(****************************************************************************************************<br>
© Syntegon Group.<br>
All rights reserved, also regarding any disposal, exploitation, reproduction, editing, distribution,<br>
as well as in the event of applications for industrial property rights.<br>
*****************************************************************************************************<br>
DESCRIPTION:<br>
Answers the waiting machine command: accepted, or rejected with the reason the Simulator shows. The command no<br>
longer waits afterwards.<br>
*****************************************************************************************************<br>
OUTPUT VALUES:<br>
FALSE while no command waits.<br>
****************************************************************************************************)
METHOD m_AnswerCommand : BOOL
VAR_INPUT
	vi_b_Accepted						: BOOL;	// TRUE: the application carries the command out
	vi_str_Reason						: STRING(80);	// why it is rejected, '' when accepted
END_VAR
m_AnswerCommand := vo_Config.stCommand.bRequested;
IF NOT m_AnswerCommand THEN
	RETURN;
END_IF
vo_Config.stCommandStatus.nHandledCommandId := vo_Config.stCommand.nCommandId;
vo_Config.stCommandStatus.eResult := SEL(vi_b_Accepted, E_ConfigCommandResult.REJECTED, E_ConfigCommandResult.ACCEPTED);
vo_Config.stCommandStatus.sMessage := SEL(vi_b_Accepted, vi_str_Reason, '');
vo_Config.stCommand.bRequested := FALSE;
END_METHOD

(****************************************************************************************************<br>
© Syntegon Group.<br>
All rights reserved, also regarding any disposal, exploitation, reproduction, editing, distribution,<br>
as well as in the event of applications for industrial property rights.<br>
*****************************************************************************************************<br>
DESCRIPTION:<br>
The machine command waiting for the application's answer (START, STOP, RESET); NONE while none waits. Answer it<br>
with m_AnswerCommand: the application alone decides whether it is carried out.<br>
****************************************************************************************************)
METHOD m_Command : E_ConfigCommand
IF vo_Config.stCommand.bRequested THEN
	m_Command := vo_Config.stCommand.eCommand;
ELSE
	m_Command := E_ConfigCommand.NONE;
END_IF
END_METHOD

(****************************************************************************************************<br>
© Syntegon Group.<br>
All rights reserved, also regarding any disposal, exploitation, reproduction, editing, distribution,<br>
as well as in the event of applications for industrial property rights.<br>
*****************************************************************************************************<br>
DESCRIPTION:<br>
Every cycle, after the fields are declared: handles a staged recipe or a reset (a recipe only while<br>
vi_b_ApplyAllowed), keeps the active recipe in vio_Set and gives the effective values in vo_Config.aActive: the<br>
active recipe while one is valid, else the fields' program values.<br>
*****************************************************************************************************<br>
OUTPUT VALUES:<br>
TRUE in the cycle a recipe was taken over or reset.<br>
****************************************************************************************************)
METHOD m_Cycle : BOOL
VAR_IN_OUT
	vio_Set								: ST_ConfigRecipeSet;	// the application's VAR PERSISTENT active recipe
END_VAR
VAR_INPUT
	vi_b_ApplyAllowed					: BOOL;	// [-] a staged recipe may be taken over now, e.g. while the machine stands
END_VAR
VAR
	str_TempRejection					: STRING(80);
	un_TempIndex						: UINT;
END_VAR
m_Cycle := FALSE;
CASE m_Staging(vio_Staging := vo_Config.stStaging, vio_Status := vo_Config.stStatus, vi_b_ApplyAllowed := vi_b_ApplyAllowed,
	vi_udn_ActiveVersion := SEL(vio_Set.bValid, 0, vio_Set.nVersion)) OF
	E_ConfigAction.RESET:
		vio_Set.bValid := FALSE;
		m_Handled(vio_Staging := vo_Config.stStaging, vio_Status := vo_Config.stStatus, vi_str_Rejection := '');
		m_Cycle := TRUE;
	E_ConfigAction.TAKE_OVER:
		str_TempRejection := m_Invalid();
		IF str_TempRejection = '' THEN
			vio_Set.nLastVersion := vio_Set.nLastVersion + 1;
			vio_Set.nVersion := vio_Set.nLastVersion;
			vio_Set.aValues := vo_Config.aStaged;
			vio_Set.bValid := TRUE;
			m_Cycle := TRUE;
		END_IF
		m_Handled(vio_Staging := vo_Config.stStaging, vio_Status := vo_Config.stStatus, vi_str_Rejection := str_TempRejection);
END_CASE


(****************************************************************************************************
EFFECTIVE VALUES
****************************************************************************************************)
un_TempIndex := 0;
WHILE un_TempIndex < vo_Config.nFieldCount AND un_TempIndex < CONFIG_GlobalConst_Param.CONFIG_un_MAX_RECIPE_FIELDS DO
	vo_Config.aActive[un_TempIndex] := SEL(vio_Set.bValid, vo_Config.aFields[un_TempIndex].fProgramValue,
		vio_Set.aValues[un_TempIndex]);
	un_TempIndex := un_TempIndex + 1;
END_WHILE
vo_Config.stStatus.nActiveVersion := SEL(vio_Set.bValid, 0, vio_Set.nVersion);
END_METHOD

(****************************************************************************************************<br>
© Syntegon Group.<br>
All rights reserved, also regarding any disposal, exploitation, reproduction, editing, distribution,<br>
as well as in the event of applications for industrial property rights.<br>
*****************************************************************************************************<br>
DESCRIPTION:<br>
Declares recipe field vi_un_Field (1..CONFIG_un_MAX_RECIPE_FIELDS): its name, the component it belongs to, how its<br>
value is kept, its unit, range and the program value that applies while no recipe is active. Fields are listed up<br>
to the highest one declared. Idempotent: call it every cycle, before m_Cycle. A CHOICE field's values are named with<br>
m_SetChoice and range from 0; its vi_lr_Min and vi_lr_Max are not used, nor a SWITCH's.<br>
*****************************************************************************************************<br>
OUTPUT VALUES:<br>
FALSE for vi_un_Field = 0 or above CONFIG_un_MAX_RECIPE_FIELDS.<br>
****************************************************************************************************)
METHOD m_DeclareField : BOOL
VAR_INPUT
	vi_un_Field							: UINT;	// [-] 1..CONFIG_un_MAX_RECIPE_FIELDS
	vi_str_Name							: STRING(31);	// unique in the recipe, e.g. 'BeltSpeed'
	vi_udn_Group						: UDINT;	// [-] manifest id of the Syn_Visu component, 0 = the whole machine
	vi_e_Type							: E_ConfigFieldType;
	vi_str_Unit							: STRING(15);	// e.g. 'mm/s', '' = none
	vi_lr_Min							: LREAL;	// smallest value of a NUMBER or INTEGER field
	vi_lr_Max							: LREAL;	// largest value of a NUMBER or INTEGER field
	vi_lr_ProgramValue					: LREAL;	// the application's own value; a SWITCH: 1 = on
END_VAR
m_DeclareField := vi_un_Field > 0 AND vi_un_Field <= CONFIG_GlobalConst_Param.CONFIG_un_MAX_RECIPE_FIELDS;
IF NOT m_DeclareField THEN
	RETURN;
END_IF
vo_Config.aFields[vi_un_Field - 1].sName := vi_str_Name;
vo_Config.aFields[vi_un_Field - 1].nGroup := vi_udn_Group;
vo_Config.aFields[vi_un_Field - 1].eType := vi_e_Type;
vo_Config.aFields[vi_un_Field - 1].sUnit := vi_str_Unit;
vo_Config.aFields[vi_un_Field - 1].fMin := vi_lr_Min;
vo_Config.aFields[vi_un_Field - 1].fMax := vi_lr_Max;
vo_Config.aFields[vi_un_Field - 1].fProgramValue := vi_lr_ProgramValue;
IF vi_un_Field > vo_Config.nFieldCount THEN
	vo_Config.nFieldCount := vi_un_Field;
END_IF
END_METHOD

(****************************************************************************************************<br>
© Syntegon Group.<br>
All rights reserved, also regarding any disposal, exploitation, reproduction, editing, distribution,<br>
as well as in the event of applications for industrial property rights.<br>
*****************************************************************************************************<br>
DESCRIPTION:<br>
Effective value of an INTEGER or CHOICE recipe field as a whole number (see m_Value).<br>
****************************************************************************************************)
METHOD m_Integer : DINT
VAR_INPUT
	vi_un_Field							: UINT;	// [-] 1..the field count
END_VAR
m_Integer := LREAL_TO_DINT(m_Value(vi_un_Field := vi_un_Field));
END_METHOD

(****************************************************************************************************<br>
© Syntegon Group.<br>
All rights reserved, also regarding any disposal, exploitation, reproduction, editing, distribution,<br>
as well as in the event of applications for industrial property rights.<br>
*****************************************************************************************************<br>
DESCRIPTION:<br>
Why the staged recipe cannot be taken over; '' when it can: a value outside its field's range (NUMBER, INTEGER),<br>
not one of its choices (CHOICE), not a whole number (INTEGER, CHOICE) or not 0 or 1 (SWITCH).<br>
****************************************************************************************************)
METHOD PRIVATE m_Invalid : STRING(80)
VAR
	un_TempIndex						: UINT;
	lr_TempValue						: LREAL;
	lr_TempMin							: LREAL;
	lr_TempMax							: LREAL;
END_VAR
m_Invalid := '';
un_TempIndex := 0;
WHILE un_TempIndex < vo_Config.nFieldCount AND un_TempIndex < CONFIG_GlobalConst_Param.CONFIG_un_MAX_RECIPE_FIELDS DO
	lr_TempValue := vo_Config.aStaged[un_TempIndex];
	CASE vo_Config.aFields[un_TempIndex].eType OF
		E_ConfigFieldType.SWITCH:
			lr_TempMin := 0;
			lr_TempMax := 1;
		E_ConfigFieldType.CHOICE:
			lr_TempMin := 0;
			lr_TempMax := UINT_TO_LREAL(vo_Config.aFields[un_TempIndex].nChoiceCount) - 1;
	ELSE
		lr_TempMin := vo_Config.aFields[un_TempIndex].fMin;
		lr_TempMax := vo_Config.aFields[un_TempIndex].fMax;
	END_CASE
	(* The range first: only a value in range is turned into a whole number. NaN equals nothing, not even itself. *)
	IF lr_TempValue <> lr_TempValue OR lr_TempValue < lr_TempMin OR lr_TempValue > lr_TempMax THEN
		m_Invalid := CONCAT(CONCAT('Field ', vo_Config.aFields[un_TempIndex].sName), CONCAT(': ', CONCAT(LREAL_TO_STRING(lr_TempValue),
			CONCAT(' is outside ', CONCAT(LREAL_TO_STRING(lr_TempMin), CONCAT(' to ', LREAL_TO_STRING(lr_TempMax)))))));
		RETURN;
	END_IF
	IF vo_Config.aFields[un_TempIndex].eType <> E_ConfigFieldType.NUMBER
		AND LINT_TO_LREAL(LREAL_TO_LINT(lr_TempValue)) <> lr_TempValue
	THEN
		m_Invalid := CONCAT(CONCAT('Field ', vo_Config.aFields[un_TempIndex].sName), CONCAT(': ',
			CONCAT(LREAL_TO_STRING(lr_TempValue), ' is not a value of its type')));
		RETURN;
	END_IF
	un_TempIndex := un_TempIndex + 1;
END_WHILE
END_METHOD

(****************************************************************************************************<br>
© Syntegon Group.<br>
All rights reserved, also regarding any disposal, exploitation, reproduction, editing, distribution,<br>
as well as in the event of applications for industrial property rights.<br>
*****************************************************************************************************<br>
DESCRIPTION:<br>
Names value vi_un_Value (0..CONFIG_un_MAX_CHOICES-1) of the CHOICE field vi_un_Field, e.g. 0 = 'Lanes'. The field<br>
has as many choices as the highest value named plus one. Idempotent: call it every cycle with m_DeclareField.<br>
*****************************************************************************************************<br>
OUTPUT VALUES:<br>
FALSE for a field not declared or a value above CONFIG_un_MAX_CHOICES - 1.<br>
****************************************************************************************************)
METHOD m_SetChoice : BOOL
VAR_INPUT
	vi_un_Field							: UINT;	// [-] the field, 1..its count
	vi_un_Value							: UINT;	// [-] the value it names, from 0
	vi_str_Text							: STRING(31);	// e.g. 'Lanes'
END_VAR
m_SetChoice := vi_un_Field > 0 AND vi_un_Field <= vo_Config.nFieldCount
	AND vi_un_Value < CONFIG_GlobalConst_Param.CONFIG_un_MAX_CHOICES;
IF NOT m_SetChoice THEN
	RETURN;
END_IF
vo_Config.aFields[vi_un_Field - 1].aChoices[vi_un_Value] := vi_str_Text;
IF vi_un_Value >= vo_Config.aFields[vi_un_Field - 1].nChoiceCount THEN
	vo_Config.aFields[vi_un_Field - 1].nChoiceCount := vi_un_Value + 1;
END_IF
END_METHOD

(****************************************************************************************************<br>
© Syntegon Group.<br>
All rights reserved, also regarding any disposal, exploitation, reproduction, editing, distribution,<br>
as well as in the event of applications for industrial property rights.<br>
*****************************************************************************************************<br>
DESCRIPTION:<br>
Gives the declared field vi_un_Field the label the Simulator shows instead of its name put into words, and a<br>
description of what it is for, shown in the field's tooltip (config protocol 4, #49). Free text in the operators'<br>
language; the name stays the field's key. Idempotent: call it every cycle with m_DeclareField.<br>
*****************************************************************************************************<br>
OUTPUT VALUES:<br>
FALSE for a field not declared.<br>
****************************************************************************************************)
METHOD m_SetText : BOOL
VAR_INPUT
	vi_un_Field							: UINT;	// [-] the field, 1..its count
	vi_str_Label						: STRING(40);	// e.g. 'Belt speed', '' = the name put into words
	vi_str_Description					: STRING(160);	// what the field is for, '' = none
END_VAR
m_SetText := vi_un_Field > 0 AND vi_un_Field <= vo_Config.nFieldCount;
IF NOT m_SetText THEN
	RETURN;
END_IF
vo_Config.aFields[vi_un_Field - 1].sLabel := vi_str_Label;
vo_Config.aFields[vi_un_Field - 1].sDescription := vi_str_Description;
END_METHOD

(****************************************************************************************************<br>
© Syntegon Group.<br>
All rights reserved, also regarding any disposal, exploitation, reproduction, editing, distribution,<br>
as well as in the event of applications for industrial property rights.<br>
*****************************************************************************************************<br>
DESCRIPTION:<br>
Shows the declared field vi_un_Field in the Simulator only while field vi_un_OnField has the value vi_dn_Value<br>
(config protocol 4, #49), e.g. a lane count only while the pattern is Lanes. vi_un_OnField must be a SWITCH (0 / 1),<br>
CHOICE or INTEGER field and may belong to another group; a field depending on a hidden one is hidden too. A hidden<br>
field keeps its value and is written with the recipe. vi_un_OnField = 0 shows the field always. The gateway reports<br>
a condition on a NUMBER field, on the field itself, on a field not declared, on a value that field can never have<br>
or in a ring as a discovery error and shows that field always. Idempotent: call it every cycle with m_DeclareField.<br>
*****************************************************************************************************<br>
OUTPUT VALUES:<br>
FALSE for a field not declared.<br>
****************************************************************************************************)
METHOD m_SetVisibleWhen : BOOL
VAR_INPUT
	vi_un_Field							: UINT;	// [-] the field shown on condition, 1..its count
	vi_un_OnField						: UINT;	// [-] the field the condition reads, 0 = always shown
	vi_dn_Value							: DINT;	// [-] the value vi_un_OnField must have
END_VAR
m_SetVisibleWhen := vi_un_Field > 0 AND vi_un_Field <= vo_Config.nFieldCount;
IF NOT m_SetVisibleWhen THEN
	RETURN;
END_IF
vo_Config.aFields[vi_un_Field - 1].nVisibleField := vi_un_OnField;
vo_Config.aFields[vi_un_Field - 1].nVisibleValue := vi_dn_Value;
END_METHOD

(****************************************************************************************************<br>
© Syntegon Group.<br>
All rights reserved, also regarding any disposal, exploitation, reproduction, editing, distribution,<br>
as well as in the event of applications for industrial property rights.<br>
*****************************************************************************************************<br>
DESCRIPTION:<br>
Effective value of a SWITCH recipe field: TRUE for on (see m_Value).<br>
****************************************************************************************************)
METHOD m_Switch : BOOL
VAR_INPUT
	vi_un_Field							: UINT;	// [-] 1..the field count
END_VAR
m_Switch := m_Value(vi_un_Field := vi_un_Field) <> 0;
END_METHOD

(****************************************************************************************************<br>
© Syntegon Group.<br>
All rights reserved, also regarding any disposal, exploitation, reproduction, editing, distribution,<br>
as well as in the event of applications for industrial property rights.<br>
*****************************************************************************************************<br>
DESCRIPTION:<br>
Effective value of recipe field vi_un_Field, for the application's logic: the active recipe's, else the program<br>
value. 0 for a field not declared. A SWITCH gives 1 or 0, an INTEGER or CHOICE a whole number (m_Switch,<br>
m_Integer give them typed).<br>
****************************************************************************************************)
METHOD m_Value : LREAL
VAR_INPUT
	vi_un_Field							: UINT;	// [-] 1..the field count
END_VAR
IF vi_un_Field > 0 AND vi_un_Field <= vo_Config.nFieldCount THEN
	m_Value := vo_Config.aActive[vi_un_Field - 1];
ELSE
	m_Value := 0;
END_IF
END_METHOD

END_FUNCTION_BLOCK

// POUs/_FB_ConfigCartesian
(****************************************************************************************************<br>
© Syntegon Group.<br>
All rights reserved, also regarding any disposal, exploitation, reproduction, editing, distribution,<br>
as well as in the event of applications for industrial property rights.<br>
*****************************************************************************************************<br>
DESCRIPTION:<br>
Parameter set of one Cartesian robot (ADR 0017): its pose, origin shift, zones, gripper fingers, limit area and<br>
TCP limit area, written by the configurator, taken over when the application allows it.<br>
Typical cycle:<br>
  fb_CartParam.m_Register(vio_Manifest := GVL_Config.stManifest, vi_udn_Id := fb_Cart.m_Id());<br>
  fb_CartParam.m_Cycle(vio_Default := CartDefault, vio_Set := CartSet, vi_b_ApplyAllowed := b_Stopped);<br>
  fb_Cart.m_Configure(vi_Pose := fb_CartParam.m_Pose(), vi_lr_XMin := 0, ...);<br>
  fb_CartParam.m_PassOn(vio_Visu := fb_Cart);<br>
The application's logic takes its zones and limit areas from m_Active, not from its own constants.<br>
*****************************************************************************************************<br>
OUTPUT VALUES:<br>
vo_Config is the contract structure the gateway reads and writes at the path in the config manifest.<br>
*****************************************************************************************************<br>
VERSION         ¦ DATE       ¦ NAME      ¦ CHANGE<br>
Syn_Config 1.1.0 ¦ 2026-11-10 ¦ J.Willner ¦ New<br>
Syn_Config 2.0.0 ¦ 2026-11-11 ¦ J.Willner ¦ Gripper fingers with their offsets, m_Invalid (ADR 0018)<br>
****************************************************************************************************)
FUNCTION_BLOCK _FB_ConfigCartesian EXTENDS _FB_ConfigComponent
VAR_OUTPUT
	vo_Config							: ST_ConfigCartesian;	// contract structure of the gateway
END_VAR

(****************************************************************************************************<br>
© Syntegon Group.<br>
All rights reserved, also regarding any disposal, exploitation, reproduction, editing, distribution,<br>
as well as in the event of applications for industrial property rights.<br>
*****************************************************************************************************<br>
DESCRIPTION:<br>
All effective values (zones, limit areas, ...), for the application's own logic.<br>
****************************************************************************************************)
METHOD m_Active : ST_ConfigCartesianParam
m_Active := vo_Config.stActive;
END_METHOD

(****************************************************************************************************<br>
© Syntegon Group.<br>
All rights reserved, also regarding any disposal, exploitation, reproduction, editing, distribution,<br>
as well as in the event of applications for industrial property rights.<br>
*****************************************************************************************************<br>
DESCRIPTION:<br>
A Cartesian robot.<br>
****************************************************************************************************)
METHOD PROTECTED m_ComponentType : SynVisu.E_VisuComponentType
m_ComponentType := SynVisu.E_VisuComponentType.CARTESIAN;
END_METHOD

(****************************************************************************************************<br>
© Syntegon Group.<br>
All rights reserved, also regarding any disposal, exploitation, reproduction, editing, distribution,<br>
as well as in the event of applications for industrial property rights.<br>
*****************************************************************************************************<br>
DESCRIPTION:<br>
Every cycle: handles a staged set or a reset (a set only while vi_b_ApplyAllowed), keeps the active set in<br>
vio_Set and gives the effective values in vo_Config.stActive: the active set while one is valid, else the<br>
program values vio_Default.<br>
*****************************************************************************************************<br>
OUTPUT VALUES:<br>
TRUE in the cycle a set was taken over or reset.<br>
****************************************************************************************************)
METHOD m_Cycle : BOOL
VAR_IN_OUT CONSTANT
	vio_Default							: ST_ConfigCartesianParam;	// the application's program values
END_VAR
VAR_IN_OUT
	vio_Set								: ST_ConfigCartesianSet;	// the application's VAR PERSISTENT active set
END_VAR
VAR_INPUT
	vi_b_ApplyAllowed					: BOOL;	// [-] a staged set may be taken over now, e.g. while the machine stands
END_VAR
VAR
	str_TempRejection					: STRING(80);
END_VAR
m_Cycle := FALSE;
CASE m_Staging(vio_Staging := vo_Config.stStaging, vio_Status := vo_Config.stStatus, vi_b_ApplyAllowed := vi_b_ApplyAllowed,
	vi_udn_ActiveVersion := SEL(vio_Set.bValid, 0, vio_Set.nVersion)) OF
	E_ConfigAction.RESET:
		vio_Set.bValid := FALSE;
		m_Handled(vio_Staging := vo_Config.stStaging, vio_Status := vo_Config.stStatus, vi_str_Rejection := '');
		m_Cycle := TRUE;
	E_ConfigAction.TAKE_OVER:
		str_TempRejection := m_Invalid(vio_Param := vo_Config.stStaged);
		IF str_TempRejection = '' THEN
			vio_Set.nLastVersion := vio_Set.nLastVersion + 1;
			vio_Set.nVersion := vio_Set.nLastVersion;
			vio_Set.stParam := vo_Config.stStaged;
			vio_Set.bValid := TRUE;
			m_Cycle := TRUE;
		END_IF
		m_Handled(vio_Staging := vo_Config.stStaging, vio_Status := vo_Config.stStatus, vi_str_Rejection := str_TempRejection);
END_CASE


(****************************************************************************************************
EFFECTIVE VALUES
****************************************************************************************************)
IF vio_Set.bValid THEN
	vo_Config.stActive := vio_Set.stParam;
	vo_Config.stStatus.nActiveVersion := vio_Set.nVersion;
ELSE
	vo_Config.stActive := vio_Default;
	vo_Config.stStatus.nActiveVersion := 0;
END_IF
END_METHOD

(****************************************************************************************************<br>
© Syntegon Group.<br>
All rights reserved, also regarding any disposal, exploitation, reproduction, editing, distribution,<br>
as well as in the event of applications for industrial property rights.<br>
*****************************************************************************************************<br>
DESCRIPTION:<br>
Why a staged set cannot be taken over; '' when it can: more zones or fingers than the lists hold, a zone on no<br>
conveyor (id 0), or a finger without a diameter or height.<br>
****************************************************************************************************)
METHOD PRIVATE m_Invalid : STRING(80)
VAR_IN_OUT CONSTANT
	vio_Param							: ST_ConfigCartesianParam;	// the staged set
END_VAR
m_Invalid := m_InvalidZones(vio_aZones := vio_Param.aZones, vi_un_Count := vio_Param.nZoneCount);
IF m_Invalid = '' THEN
	m_Invalid := m_InvalidFingers(vio_aFingers := vio_Param.aFingers, vi_un_Count := vio_Param.nFingerCount);
END_IF
END_METHOD

(****************************************************************************************************<br>
© Syntegon Group.<br>
All rights reserved, also regarding any disposal, exploitation, reproduction, editing, distribution,<br>
as well as in the event of applications for industrial property rights.<br>
*****************************************************************************************************<br>
DESCRIPTION:<br>
Passes the effective origin shift, limit areas, zones and fingers on to the robot's Syn_Visu FB, so the<br>
visualisation shows what the machine uses. The pose goes with the application's own m_Configure call (with<br>
the strokes and rail height, hardware): vi_Pose := m_Pose(). Call it after m_Cycle, every cycle; Syn_Visu's<br>
config version only changes when a value does.<br>
****************************************************************************************************)
METHOD m_PassOn : BOOL
VAR_IN_OUT
	vio_Visu							: SynVisu._FB_VisuCartesian;	// the robot's Syn_Visu FB
END_VAR
m_PassOn := TRUE;
vio_Visu.m_SetOriginShift(vi_lr_X := vo_Config.stActive.stOriginShift.fX, vi_lr_Y := vo_Config.stActive.stOriginShift.fY,
	vi_lr_Z := vo_Config.stActive.stOriginShift.fZ);
m_PassOnLimitAreas(vio_Visu := vio_Visu, vio_LimitArea := vo_Config.stActive.stLimitArea,
	vio_TcpLimitArea := vo_Config.stActive.stTcpLimitArea);
m_PassOnZones(vio_Visu := vio_Visu, vio_aZones := vo_Config.stActive.aZones, vi_un_Count := vo_Config.stActive.nZoneCount,
	vi_un_VisuCount := vio_Visu.vo_Visu.stConfig.nZoneCount);
m_PassOnFingers(vio_Visu := vio_Visu, vio_aFingers := vo_Config.stActive.aFingers,
	vi_un_Count := vo_Config.stActive.nFingerCount, vi_un_VisuCount := vio_Visu.vo_Visu.stConfig.nFingerCount);
END_METHOD

(****************************************************************************************************<br>
© Syntegon Group.<br>
All rights reserved, also regarding any disposal, exploitation, reproduction, editing, distribution,<br>
as well as in the event of applications for industrial property rights.<br>
*****************************************************************************************************<br>
DESCRIPTION:<br>
Effective pose of the axis origin (MCS), for the application's logic and its Syn_Visu m_Configure call.<br>
****************************************************************************************************)
METHOD m_Pose : SynVisu.ST_VisuPose
m_Pose := vo_Config.stActive.stPose;
END_METHOD

END_FUNCTION_BLOCK

// POUs/_FB_ConfigXtsLoop
(****************************************************************************************************<br>
© Syntegon Group.<br>
All rights reserved, also regarding any disposal, exploitation, reproduction, editing, distribution,<br>
as well as in the event of applications for industrial property rights.<br>
*****************************************************************************************************<br>
DESCRIPTION:<br>
Parameter set of one XTS loop (ADR 0017): its pose, origin shift, track modules, zones and gripper fingers,<br>
written by the configurator, taken over when the application allows it. Typical cycle:<br>
  fb_FxxParam.m_Register(vio_Manifest := GVL_Config.stManifest, vi_udn_Id := fb_Fxx.m_Id());<br>
  fb_FxxParam.m_Cycle(vio_Default := FxxDefault, vio_Set := FxxSet, vi_b_ApplyAllowed := b_Stopped);<br>
  fb_Fxx.m_Configure(vi_Pose := fb_FxxParam.m_Pose(), vi_lr_ToolOffset := 120, ...);<br>
  fb_FxxParam.m_PassOn(vio_Visu := fb_Fxx);<br>
The application's logic takes its track and zones from m_Active, not from its own constants.<br>
*****************************************************************************************************<br>
OUTPUT VALUES:<br>
vo_Config is the contract structure the gateway reads and writes at the path in the config manifest.<br>
*****************************************************************************************************<br>
VERSION         ¦ DATE       ¦ NAME      ¦ CHANGE<br>
Syn_Config 1.1.0 ¦ 2026-11-10 ¦ J.Willner ¦ New<br>
Syn_Config 2.0.0 ¦ 2026-11-11 ¦ J.Willner ¦ Gripper fingers with their offsets (ADR 0018)<br>
****************************************************************************************************)
FUNCTION_BLOCK _FB_ConfigXtsLoop EXTENDS _FB_ConfigComponent
VAR_OUTPUT
	vo_Config							: ST_ConfigXtsLoop;	// contract structure of the gateway
END_VAR

(****************************************************************************************************<br>
© Syntegon Group.<br>
All rights reserved, also regarding any disposal, exploitation, reproduction, editing, distribution,<br>
as well as in the event of applications for industrial property rights.<br>
*****************************************************************************************************<br>
DESCRIPTION:<br>
All effective values (track modules, zones, ...), for the application's own logic.<br>
****************************************************************************************************)
METHOD m_Active : ST_ConfigXtsLoopParam
m_Active := vo_Config.stActive;
END_METHOD

(****************************************************************************************************<br>
© Syntegon Group.<br>
All rights reserved, also regarding any disposal, exploitation, reproduction, editing, distribution,<br>
as well as in the event of applications for industrial property rights.<br>
*****************************************************************************************************<br>
DESCRIPTION:<br>
An XTS loop.<br>
****************************************************************************************************)
METHOD PROTECTED m_ComponentType : SynVisu.E_VisuComponentType
m_ComponentType := SynVisu.E_VisuComponentType.XTS_LOOP;
END_METHOD

(****************************************************************************************************<br>
© Syntegon Group.<br>
All rights reserved, also regarding any disposal, exploitation, reproduction, editing, distribution,<br>
as well as in the event of applications for industrial property rights.<br>
*****************************************************************************************************<br>
DESCRIPTION:<br>
Every cycle: handles a staged set or a reset (a set only while vi_b_ApplyAllowed), keeps the active set in<br>
vio_Set and gives the effective values in vo_Config.stActive: the active set while one is valid, else the<br>
program values vio_Default.<br>
*****************************************************************************************************<br>
OUTPUT VALUES:<br>
TRUE in the cycle a set was taken over or reset.<br>
****************************************************************************************************)
METHOD m_Cycle : BOOL
VAR_IN_OUT CONSTANT
	vio_Default							: ST_ConfigXtsLoopParam;	// the application's program values
END_VAR
VAR_IN_OUT
	vio_Set								: ST_ConfigXtsLoopSet;	// the application's VAR PERSISTENT active set
END_VAR
VAR_INPUT
	vi_b_ApplyAllowed					: BOOL;	// [-] a staged set may be taken over now, e.g. while the machine stands
END_VAR
VAR
	str_TempRejection					: STRING(80);
END_VAR
m_Cycle := FALSE;
CASE m_Staging(vio_Staging := vo_Config.stStaging, vio_Status := vo_Config.stStatus, vi_b_ApplyAllowed := vi_b_ApplyAllowed,
	vi_udn_ActiveVersion := SEL(vio_Set.bValid, 0, vio_Set.nVersion)) OF
	E_ConfigAction.RESET:
		vio_Set.bValid := FALSE;
		m_Handled(vio_Staging := vo_Config.stStaging, vio_Status := vo_Config.stStatus, vi_str_Rejection := '');
		m_Cycle := TRUE;
	E_ConfigAction.TAKE_OVER:
		str_TempRejection := m_Invalid(vio_Param := vo_Config.stStaged);
		IF str_TempRejection = '' THEN
			vio_Set.nLastVersion := vio_Set.nLastVersion + 1;
			vio_Set.nVersion := vio_Set.nLastVersion;
			vio_Set.stParam := vo_Config.stStaged;
			vio_Set.bValid := TRUE;
			m_Cycle := TRUE;
		END_IF
		m_Handled(vio_Staging := vo_Config.stStaging, vio_Status := vo_Config.stStatus, vi_str_Rejection := str_TempRejection);
END_CASE


(****************************************************************************************************
EFFECTIVE VALUES
****************************************************************************************************)
IF vio_Set.bValid THEN
	vo_Config.stActive := vio_Set.stParam;
	vo_Config.stStatus.nActiveVersion := vio_Set.nVersion;
ELSE
	vo_Config.stActive := vio_Default;
	vo_Config.stStatus.nActiveVersion := 0;
END_IF
END_METHOD

(****************************************************************************************************<br>
© Syntegon Group.<br>
All rights reserved, also regarding any disposal, exploitation, reproduction, editing, distribution,<br>
as well as in the event of applications for industrial property rights.<br>
*****************************************************************************************************<br>
DESCRIPTION:<br>
Why a staged set cannot be taken over; '' when it can: a track without modules, more modules, zones or fingers<br>
than the lists hold, a module without a length, a zone on no conveyor (id 0), or a finger without a diameter or<br>
height.<br>
****************************************************************************************************)
METHOD PRIVATE m_Invalid : STRING(80)
VAR_IN_OUT CONSTANT
	vio_Param							: ST_ConfigXtsLoopParam;	// the staged set
END_VAR
m_Invalid := m_InvalidModules(vio_aModules := vio_Param.aModules, vi_un_Count := vio_Param.nModuleCount);
IF m_Invalid = '' THEN
	m_Invalid := m_InvalidZones(vio_aZones := vio_Param.aZones, vi_un_Count := vio_Param.nZoneCount);
END_IF
IF m_Invalid = '' THEN
	m_Invalid := m_InvalidFingers(vio_aFingers := vio_Param.aFingers, vi_un_Count := vio_Param.nFingerCount);
END_IF
END_METHOD

(****************************************************************************************************<br>
© Syntegon Group.<br>
All rights reserved, also regarding any disposal, exploitation, reproduction, editing, distribution,<br>
as well as in the event of applications for industrial property rights.<br>
*****************************************************************************************************<br>
DESCRIPTION:<br>
Passes the effective origin shift, track modules, zones and fingers on to the loop's Syn_Visu FB, so the<br>
visualisation shows what the machine uses. The pose goes with the application's own m_Configure call (with<br>
the tool offset and mover size, hardware): vi_Pose := m_Pose(). Call it after m_Cycle, every cycle; Syn_Visu's<br>
config version only changes when a value does.<br>
****************************************************************************************************)
METHOD m_PassOn : BOOL
VAR_IN_OUT
	vio_Visu							: SynVisu._FB_VisuXtsLoop;	// the loop's Syn_Visu FB
END_VAR
m_PassOn := TRUE;
vio_Visu.m_SetOriginShift(vi_lr_X := vo_Config.stActive.stOriginShift.fX, vi_lr_Y := vo_Config.stActive.stOriginShift.fY,
	vi_lr_Z := vo_Config.stActive.stOriginShift.fZ);
m_PassOnModules(vio_Visu := vio_Visu, vio_aModules := vo_Config.stActive.aModules,
	vi_un_Count := vo_Config.stActive.nModuleCount, vi_un_VisuCount := vio_Visu.vo_Visu.stConfig.nModuleCount);
m_PassOnZones(vio_Visu := vio_Visu, vio_aZones := vo_Config.stActive.aZones, vi_un_Count := vo_Config.stActive.nZoneCount,
	vi_un_VisuCount := vio_Visu.vo_Visu.stConfig.nZoneCount);
m_PassOnFingers(vio_Visu := vio_Visu, vio_aFingers := vo_Config.stActive.aFingers,
	vi_un_Count := vo_Config.stActive.nFingerCount, vi_un_VisuCount := vio_Visu.vo_Visu.stConfig.nFingerCount);
END_METHOD

(****************************************************************************************************<br>
© Syntegon Group.<br>
All rights reserved, also regarding any disposal, exploitation, reproduction, editing, distribution,<br>
as well as in the event of applications for industrial property rights.<br>
*****************************************************************************************************<br>
DESCRIPTION:<br>
Effective pose of the start of module 1 (MCS), for the application's logic and its Syn_Visu m_Configure call.<br>
****************************************************************************************************)
METHOD m_Pose : SynVisu.ST_VisuPose
m_Pose := vo_Config.stActive.stPose;
END_METHOD

END_FUNCTION_BLOCK

// POUs/_FC_GetVersionSynConfig
(****************************************************************************************************<br>
© Syntegon Group.<br>
All rights reserved, also regarding any disposal, exploitation, reproduction, editing, distribution,<br>
as well as in the event of applications for industrial property rights.<br>
*****************************************************************************************************<br>
DESCRIPTION:<br>
Runtime-readable version of the Syn_Config library.<br>
*****************************************************************************************************<br>
VERSION         ¦ DATE       ¦ NAME      ¦ CHANGE<br>
Syn_Config 1.0.0 ¦ 2026-11-10 ¦ J.Willner ¦ Parameter sets of conveyors and Deltas (ADR 0017, protocol 1)<br>
Syn_Config 1.1.0 ¦ 2026-11-10 ¦ J.Willner ¦ Every other component type (#24)<br>
Syn_Config 2.0.0 ¦ 2026-11-11 ¦ J.Willner ¦ Gripper fingers in the robots' sets (protocol 2, #25)<br>
Syn_Config 2.0.1 ¦ 2026-11-12 ¦ J.Willner ¦ SynVisu as a placeholder: the application chooses its version<br>
Syn_Config 2.1.0 ¦ 2026-11-14 ¦ J.Willner ¦ Machine FB: recipe fields and machine commands (protocol 3, #43)<br>
Syn_Config 2.2.0 ¦ 2026-11-14 ¦ J.Willner ¦ Recipe fields: label, description, visibility condition (protocol 4, #49)<br>
****************************************************************************************************)
FUNCTION _FC_GetVersionSynConfig : UINT
VAR_INPUT
	vi_n_VersionElement					: INT;	// [-] 1 = major, 2 = minor, 3 = revision
END_VAR

CASE vi_n_VersionElement OF
	1: _FC_GetVersionSynConfig := 2;
	2: _FC_GetVersionSynConfig := 2;
	3: _FC_GetVersionSynConfig := 0;
ELSE
	_FC_GetVersionSynConfig := 16#FFFF;
END_CASE

END_FUNCTION
